   #r := FALSE;
   #a1 := W#16#0000;
   #a2 := W#16#0000;
   #activeDataBlock := 0;
   // PB4, STEP 5 network 1
   #a2 := #a1;
   #a1 := "ROLL_GetM"(FirstByte := 239, Width := 8);
   #a2 := #a1;
   #a1 := W#16#001E;
   #comparisonResults[0] := (WORD_TO_INT(#a2) = WORD_TO_INT(#a1));
   #r := #comparisonResults[0];
   "ROLL_State".M[23, 5] := #r;
   // PB4, STEP 5 network 2
   #a2 := #a1;
   #a1 := "ROLL_GetM"(FirstByte := 239, Width := 8);
   #a2 := #a1;
   #a1 := W#16#001F;
   #comparisonResults[1] := (WORD_TO_INT(#a2) = WORD_TO_INT(#a1));
   #r := #comparisonResults[1];
   "ROLL_State".M[23, 6] := #r;
   // PB4, STEP 5 network 3
   #a2 := #a1;
   #a1 := "ROLL_GetM"(FirstByte := 239, Width := 8);
   #a2 := #a1;
   #a1 := W#16#0023;
   #comparisonResults[2] := (WORD_TO_INT(#a2) = WORD_TO_INT(#a1));
   #r := #comparisonResults[2];
   "ROLL_State".M[24, 0] := #r;
   // PB4, STEP 5 network 4
   #a2 := #a1;
   #a1 := "ROLL_GetM"(FirstByte := 239, Width := 8);
   #a2 := #a1;
   #a1 := W#16#0024;
   #comparisonResults[3] := (WORD_TO_INT(#a2) = WORD_TO_INT(#a1));
   #r := #comparisonResults[3];
   "ROLL_State".M[24, 1] := #r;
   // PB4, STEP 5 network 5
   #a2 := #a1;
   #a1 := "ROLL_GetM"(FirstByte := 239, Width := 8);
   #a2 := #a1;
   #a1 := W#16#0025;
   #comparisonResults[4] := (WORD_TO_INT(#a2) = WORD_TO_INT(#a1));
   #r := #comparisonResults[4];
   "ROLL_State".M[24, 2] := #r;
   // PB4, STEP 5 network 6
   #a2 := #a1;
   #a1 := "ROLL_GetM"(FirstByte := 239, Width := 8);
   #a2 := #a1;
   #a1 := W#16#0026;
   #comparisonResults[5] := (WORD_TO_INT(#a2) = WORD_TO_INT(#a1));
   #r := #comparisonResults[5];
   "ROLL_State".M[24, 3] := #r;
   // PB4, STEP 5 network 7
   #a2 := #a1;
   #a1 := "ROLL_GetM"(FirstByte := 239, Width := 8);
   #a2 := #a1;
   #a1 := W#16#0027;
   #comparisonResults[6] := (WORD_TO_INT(#a2) = WORD_TO_INT(#a1));
   #r := #comparisonResults[6];
   "ROLL_State".M[24, 4] := #r;
   // PB4, STEP 5 network 8
   #a2 := #a1;
   #a1 := "ROLL_GetM"(FirstByte := 239, Width := 8);
   #a2 := #a1;
   #a1 := W#16#0032;
   #comparisonResults[7] := (WORD_TO_INT(#a2) = WORD_TO_INT(#a1));
   #r := #comparisonResults[7];
   "ROLL_State".M[25, 0] := #r;
   // PB4, STEP 5 network 9
   #a2 := #a1;
   #a1 := "ROLL_GetM"(FirstByte := 239, Width := 8);
   #a2 := #a1;
   #a1 := W#16#0033;
   #comparisonResults[8] := (WORD_TO_INT(#a2) = WORD_TO_INT(#a1));
   #r := #comparisonResults[8];
   "ROLL_State".M[25, 1] := #r;
   // PB4, STEP 5 network 10
   #a2 := #a1;
   #a1 := "ROLL_GetM"(FirstByte := 239, Width := 8);
   #a2 := #a1;
   #a1 := W#16#0034;
   #comparisonResults[9] := (WORD_TO_INT(#a2) = WORD_TO_INT(#a1));
   #r := #comparisonResults[9];
   "ROLL_State".M[25, 2] := #r;
   // PB4, STEP 5 network 11
   #a2 := #a1;
   #a1 := "ROLL_GetM"(FirstByte := 239, Width := 8);
   #a2 := #a1;
   #a1 := W#16#0035;
   #comparisonResults[10] := (WORD_TO_INT(#a2) = WORD_TO_INT(#a1));
   #r := #comparisonResults[10];
   "ROLL_State".M[25, 3] := #r;
   // PB4, STEP 5 network 12
   #a2 := #a1;
   #a1 := "ROLL_GetM"(FirstByte := 239, Width := 8);
   #a2 := #a1;
   #a1 := W#16#0037;
   #comparisonResults[11] := (WORD_TO_INT(#a2) = WORD_TO_INT(#a1));
   #r := #comparisonResults[11];
   "ROLL_State".M[25, 4] := #r;
   // PB4, STEP 5 network 13
   #a2 := #a1;
   #a1 := "ROLL_GetM"(FirstByte := 239, Width := 8);
   #a2 := #a1;
   #a1 := W#16#0038;
   #comparisonResults[12] := (WORD_TO_INT(#a2) = WORD_TO_INT(#a1));
   #r := #comparisonResults[12];
   "ROLL_State".M[25, 5] := #r;
   // PB4, STEP 5 network 14
   #a2 := #a1;
   #a1 := "ROLL_GetM"(FirstByte := 239, Width := 8);
   #a2 := #a1;
   #a1 := W#16#0039;
   #comparisonResults[13] := (WORD_TO_INT(#a2) = WORD_TO_INT(#a1));
   #r := #comparisonResults[13];
   "ROLL_State".M[25, 6] := #r;
   // PB4, STEP 5 network 15
   #a2 := #a1;
   #a1 := "ROLL_GetM"(FirstByte := 239, Width := 8);
   #a2 := #a1;
   #a1 := W#16#003A;
   #comparisonResults[14] := (WORD_TO_INT(#a2) = WORD_TO_INT(#a1));
   #r := #comparisonResults[14];
   "ROLL_State".M[25, 7] := #r;
   // PB4, STEP 5 network 16
   #a2 := #a1;
   #a1 := "ROLL_GetM"(FirstByte := 239, Width := 8);
   #a2 := #a1;
   #a1 := W#16#003C;
   #comparisonResults[15] := (WORD_TO_INT(#a2) = WORD_TO_INT(#a1));
   #r := #comparisonResults[15];
   "ROLL_State".M[26, 0] := #r;
   // PB4, STEP 5 network 17
   #a2 := #a1;
   #a1 := "ROLL_GetM"(FirstByte := 239, Width := 8);
   #a2 := #a1;
   #a1 := W#16#003D;
   #comparisonResults[16] := (WORD_TO_INT(#a2) = WORD_TO_INT(#a1));
   #r := #comparisonResults[16];
   "ROLL_State".M[26, 1] := #r;
   // PB4, STEP 5 network 18
   #a2 := #a1;
   #a1 := "ROLL_GetM"(FirstByte := 239, Width := 8);
   #a2 := #a1;
   #a1 := W#16#003E;
   #comparisonResults[17] := (WORD_TO_INT(#a2) = WORD_TO_INT(#a1));
   #r := #comparisonResults[17];
   "ROLL_State".M[26, 2] := #r;
   // PB4, STEP 5 network 19
   #a2 := #a1;
   #a1 := "ROLL_GetM"(FirstByte := 239, Width := 8);
   #a2 := #a1;
   #a1 := W#16#003F;
   #comparisonResults[18] := (WORD_TO_INT(#a2) = WORD_TO_INT(#a1));
   #r := #comparisonResults[18];
   "ROLL_State".M[26, 3] := #r;
   // PB4, STEP 5 network 20
   #a2 := #a1;
   #a1 := "ROLL_GetM"(FirstByte := 239, Width := 8);
   #a2 := #a1;
   #a1 := W#16#0041;
   #comparisonResults[19] := (WORD_TO_INT(#a2) = WORD_TO_INT(#a1));
   #r := #comparisonResults[19];
   "ROLL_State".M[26, 5] := #r;
   // PB4, STEP 5 network 21
   #a2 := #a1;
   #a1 := "ROLL_GetM"(FirstByte := 239, Width := 8);
   #a2 := #a1;
   #a1 := W#16#0042;
   #comparisonResults[20] := (WORD_TO_INT(#a2) = WORD_TO_INT(#a1));
   #r := #comparisonResults[20];
   "ROLL_State".M[26, 6] := #r;
   // PB4, STEP 5 network 22
   #a2 := #a1;
   #a1 := "ROLL_GetM"(FirstByte := 239, Width := 8);
   #a2 := #a1;
   #a1 := W#16#0045;
   #comparisonResults[21] := (WORD_TO_INT(#a2) = WORD_TO_INT(#a1));
   #r := #comparisonResults[21];
   "ROLL_State".M[27, 1] := #r;
   // PB4, STEP 5 network 23
   #a2 := #a1;
   #a1 := "ROLL_GetM"(FirstByte := 239, Width := 8);
   #a2 := #a1;
   #a1 := W#16#0048;
   #comparisonResults[22] := (WORD_TO_INT(#a2) = WORD_TO_INT(#a1));
   #r := #comparisonResults[22];
   "ROLL_State".M[27, 4] := #r;
   // PB4, STEP 5 network 24
   #a2 := #a1;
   #a1 := "ROLL_GetM"(FirstByte := 239, Width := 8);
   #a2 := #a1;
   #a1 := W#16#0049;
   #comparisonResults[23] := (WORD_TO_INT(#a2) = WORD_TO_INT(#a1));
   #r := #comparisonResults[23];
   "ROLL_State".M[27, 5] := #r;
   // PB4, STEP 5 network 25
   #a2 := #a1;
   #a1 := "ROLL_GetM"(FirstByte := 239, Width := 8);
   #a2 := #a1;
   #a1 := W#16#0063;
   #comparisonResults[24] := (WORD_TO_INT(#a2) = WORD_TO_INT(#a1));
   #r := #comparisonResults[24];
   "ROLL_State".M[27, 7] := #r;
   // PB4, STEP 5 network 26
   RETURN;
END_FUNCTION

FUNCTION "ROLL_PB50" : Void   // FC33, SCL
{ S7_Optimized_Access := 'TRUE' }
VERSION : 0.1
// stored: AutoNumber true, IsIECCheckEnabled false, SetENOAutomatically false, UDAEnableTagReadback false
   VAR_TEMP
      r : Bool;
      a1 : Word;
      a2 : Word;
      activeDataBlock : Int;
      comparisonResults : Array[0..0] of Bool;
   END_VAR
BEGIN

   #r := FALSE;
   #a1 := W#16#0000;
   #a2 := W#16#0000;
   #activeDataBlock := 0;
   // PB50, STEP 5 network 1
   #activeDataBlock := 15;
   // PB50, STEP 5 network 2
   #r := "ROLL_State".M[0, 1];
   IF #r THEN
       "ROLL_State".M[0, 2] := FALSE;
   END_IF;
   // PB50, STEP 5 network 3
   #a2 := #a1;
   #a1 := W#16#2008;
   #r := ((NOT "ROLL_State".M[0, 1]) AND "ROLL_IO".Input[3, 0]);
   "ROLL_TimerOp"(Number := 11,
                  Operation := 0,
                  Signal := #r,
                  Preset := #a1);
   // PB50, STEP 5 network 4
   #a2 := #a1;
   #a1 := W#16#1020;
   #r := "ROLL_State".M[29, 0];
   "ROLL_TimerOp"(Number := 13,
                  Operation := 0,
                  Signal := #r,
                  Preset := #a1);
   // PB50, STEP 5 network 5
   RETURN;
END_FUNCTION

FUNCTION "ROLL_PB51" : Void   // FC34, SCL
{ S7_Optimized_Access := 'TRUE' }
VERSION : 0.1
// stored: AutoNumber true, IsIECCheckEnabled false, SetENOAutomatically false, UDAEnableTagReadback false
   VAR_TEMP
      r : Bool;
      a1 : Word;
      a2 : Word;
      activeDataBlock : Int;
      comparisonResults : Array[0..0] of Bool;
   END_VAR
BEGIN

   #r := FALSE;
   #a1 := W#16#0000;
   #a2 := W#16#0000;
   #activeDataBlock := 0;
   // PB51, STEP 5 network 1
   #a2 := #a1;
   #a1 := W#16#2060;
   #r := "ROLL_IO".Output[24, 0];
   "ROLL_TimerOp"(Number := 15,
                  Operation := 0,
                  Signal := #r,
                  Preset := #a1);
   // PB51, STEP 5 network 2
   #a2 := #a1;
   #a1 := W#16#3360;
   #r := ((NOT "ROLL_IO".Input[5, 6]) AND "ROLL_State".M[31, 5]);
   "ROLL_TimerOp"(Number := 16,
                  Operation := 0,
                  Signal := #r,
                  Preset := #a1);
   // PB51, STEP 5 network 3
   #a2 := #a1;
   #a1 := W#16#1010;
   #r := "ROLL_State".M[37, 5];
   "ROLL_TimerOp"(Number := 18,
                  Operation := 0,
                  Signal := #r,
                  Preset := #a1);
   // PB51, STEP 5 network 4
   #a2 := #a1;
   #a1 := W#16#2015;
   #r := (((NOT "ROLL_IO".Input[124, 1]) AND "ROLL_IO".Output[112, 1]) OR ((NOT "ROLL_IO".Input[124, 2]) AND "ROLL_IO".Output[112, 2]));
   "ROLL_TimerOp"(Number := 19,
                  Operation := 0,
                  Signal := #r,
                  Preset := #a1);
   // PB51, STEP 5 network 5
   #a2 := #a1;
   #a1 := W#16#1010;
   #r := (("ROLL_IO".Input[123, 4] OR "ROLL_IO".Input[123, 5]) AND "ROLL_IO".Output[112, 0]);
   "ROLL_TimerOp"(Number := 20,
                  Operation := 0,
                  Signal := #r,
                  Preset := #a1);
   // PB51, STEP 5 network 6
   #a2 := #a1;
   #a1 := W#16#1050;
   #r := "ROLL_IO".Input[123, 4];
   "ROLL_TimerOp"(Number := 21,
                  Operation := 0,
                  Signal := #r,
                  Preset := #a1);
   // PB51, STEP 5 network 7
   #a2 := #a1;
   #a1 := W#16#2005;
   #r := ("ROLL_IO".Input[125, 0] AND "ROLL_IO".Input[125, 1]);
   "ROLL_TimerOp"(Number := 95,
                  Operation := 0,
                  Signal := #r,
                  Preset := #a1);
   // PB51, STEP 5 network 8
   RETURN;
END_FUNCTION

FUNCTION "ROLL_PB52" : Void   // FC35, SCL
{ S7_Optimized_Access := 'TRUE' }
VERSION : 0.1
// stored: AutoNumber true, IsIECCheckEnabled false, SetENOAutomatically false, UDAEnableTagReadback false
   VAR_TEMP
      r : Bool;
      a1 : Word;
      a2 : Word;
      activeDataBlock : Int;
      comparisonResults : Array[0..0] of Bool;
   END_VAR
BEGIN

   #r := FALSE;
   #a1 := W#16#0000;
   #a2 := W#16#0000;
   #activeDataBlock := 0;
   // PB52, STEP 5 network 1
   #activeDataBlock := 15;
   // PB52, STEP 5 network 2
   #a2 := #a1;
   #a1 := "ROLL_GetDW"(DbNumber := #activeDataBlock, Index := 17);
   #r := ((NOT "ROLL_IO".Input[5, 5]) AND (NOT "ROLL_State".M[6, 3]) AND "ROLL_IO".Input[3, 1] AND "ROLL_State".M[4, 1] AND "ROLL_State".M[40, 5]);
   "ROLL_TimerOp"(Number := 17,
                  Operation := 0,
                  Signal := #r,
                  Preset := #a1);
   // PB52, STEP 5 network 3
   #a2 := #a1;
   #a1 := "ROLL_GetDW"(DbNumber := #activeDataBlock, Index := 31);
   #r := ((NOT "ROLL_IO".Input[5, 3]) AND (NOT "ROLL_State".M[6, 1]) AND "ROLL_IO".Input[3, 1] AND "ROLL_State".M[4, 1]);
   "ROLL_TimerOp"(Number := 31,
                  Operation := 0,
                  Signal := #r,
                  Preset := #a1);
   // PB52, STEP 5 network 4
   #a2 := #a1;
   #a1 := "ROLL_GetDW"(DbNumber := #activeDataBlock, Index := 32);
   #r := ((NOT "ROLL_IO".Input[6, 0]) AND (NOT "ROLL_State".M[6, 4]) AND "ROLL_IO".Input[3, 1] AND "ROLL_State".M[4, 1]);
   "ROLL_TimerOp"(Number := 32,
                  Operation := 0,
                  Signal := #r,
                  Preset := #a1);
   // PB52, STEP 5 network 5
   #a2 := #a1;
   #a1 := "ROLL_GetDW"(DbNumber := #activeDataBlock, Index := 33);
   #r := ((NOT "ROLL_IO".Input[6, 2]) AND (NOT "ROLL_State".M[6, 5]) AND "ROLL_IO".Input[3, 1] AND "ROLL_State".M[4, 1]);
   "ROLL_TimerOp"(Number := 33,
                  Operation := 0,
                  Signal := #r,
                  Preset := #a1);
   // PB52, STEP 5 network 6
   #a2 := #a1;
   #a1 := W#16#3030;
   #r := ((NOT "ROLL_State".M[0, 4]) AND (NOT "ROLL_State".M[6, 7]) AND "ROLL_IO".Input[3, 1] AND "ROLL_State".M[4, 1]);
   "ROLL_TimerOp"(Number := 35,
                  Operation := 0,
                  Signal := #r,
                  Preset := #a1);
   // PB52, STEP 5 network 7
   #a2 := #a1;
   #a1 := W#16#3030;
   #r := ((NOT "ROLL_State".M[0, 4]) AND (NOT "ROLL_State".M[7, 0]) AND "ROLL_IO".Input[3, 1] AND "ROLL_State".M[4, 1]);
   "ROLL_TimerOp"(Number := 36,
                  Operation := 0,
                  Signal := #r,
                  Preset := #a1);
   // PB52, STEP 5 network 8
   #a2 := #a1;
   #a1 := W#16#3030;
   #r := ((NOT "ROLL_State".M[0, 4]) AND (NOT "ROLL_State".M[7, 1]) AND "ROLL_IO".Input[3, 1] AND "ROLL_State".M[4, 1]);
   "ROLL_TimerOp"(Number := 37,
                  Operation := 0,
                  Signal := #r,
                  Preset := #a1);
   // PB52, STEP 5 network 9
   #a2 := #a1;
   #a1 := W#16#3030;
   #r := ((NOT "ROLL_State".M[0, 4]) AND (NOT "ROLL_State".M[7, 2]) AND "ROLL_IO".Input[3, 1] AND "ROLL_State".M[4, 1]);
   "ROLL_TimerOp"(Number := 38,
                  Operation := 0,
                  Signal := #r,
                  Preset := #a1);
   // PB52, STEP 5 network 10
   #a2 := #a1;
   #a1 := W#16#1005;
   #r := "ROLL_IO".Input[123, 1];
   "ROLL_TimerOp"(Number := 45,
                  Operation := 0,
                  Signal := #r,
                  Preset := #a1);
   // PB52, STEP 5 network 11
   #a2 := #a1;
   #a1 := "ROLL_GetDW"(DbNumber := #activeDataBlock, Index := 58);
   #r := ("ROLL_IO".Input[3, 1] AND "ROLL_State".M[3, 6]);
   "ROLL_TimerOp"(Number := 58,
                  Operation := 1,
                  Signal := #r,
                  Preset := #a1);
   #a2 := #a1;
   #a1 := "ROLL_GetDW"(DbNumber := #activeDataBlock, Index := 59);
   #r := ("ROLL_State".M[3, 6] AND "ROLL_State".S5Timers[58].Q);
   "ROLL_TimerOp"(Number := 59,
                  Operation := 1,
                  Signal := #r,
                  Preset := #a1);
   // PB52, STEP 5 network 12
   #a2 := #a1;
   #a1 := "ROLL_GetDW"(DbNumber := #activeDataBlock, Index := 63);
   #r := (NOT "ROLL_State".S5Timers[62].Q);
   "ROLL_TimerOp"(Number := 63,
                  Operation := 0,
                  Signal := #r,
                  Preset := #a1);
   #a2 := #a1;
   #a1 := "ROLL_GetDW"(DbNumber := #activeDataBlock, Index := 62);
   #r := "ROLL_State".S5Timers[63].Q;
   "ROLL_TimerOp"(Number := 62,
                  Operation := 1,
                  Signal := #r,
                  Preset := #a1);
   #r := ((NOT "ROLL_State".M[103, 0]) AND (NOT "ROLL_State".M[103, 3]) AND (NOT "ROLL_State".M[103, 4]) AND (NOT "ROLL_State".S5Timers[119].Q));
   "ROLL_TimerOp"(Number := 62,
                  Operation := 2,
                  Signal := #r,
                  Preset := #a1);
   // PB52, STEP 5 network 13
   #a2 := #a1;
   #a1 := W#16#2010;
   #r := "ROLL_IO".Input[5, 3];
   "ROLL_TimerOp"(Number := 70,
                  Operation := 1,
                  Signal := #r,
                  Preset := #a1);
   // PB52, STEP 5 network 14
   #a2 := #a1;
   #a1 := W#16#2010;
   #r := "ROLL_IO".Input[6, 2];
   "ROLL_TimerOp"(Number := 72,
                  Operation := 1,
                  Signal := #r,
                  Preset := #a1);
   // PB52, STEP 5 network 15
   #a2 := #a1;
   #a1 := "ROLL_GetDW"(DbNumber := #activeDataBlock, Index := 85);
   #r := "ROLL_State".M[41, 0];
   "ROLL_TimerOp"(Number := 85,
                  Operation := 1,
                  Signal := #r,
                  Preset := #a1);
   // PB52, STEP 5 network 16
   RETURN;
END_FUNCTION

FUNCTION "ROLL_PB7" : Void   // FC17, SCL
{ S7_Optimized_Access := 'TRUE' }
VERSION : 0.1
// stored: AutoNumber true, IsIECCheckEnabled false, SetENOAutomatically false, UDAEnableTagReadback false
   VAR_TEMP
      r : Bool;
      a1 : Word;
      a2 : Word;
      activeDataBlock : Int;
      comparisonResults : Array[0..0] of Bool;
   END_VAR
BEGIN

   #r := FALSE;
   #a1 := W#16#0000;
   #a2 := W#16#0000;
   #activeDataBlock := 0;
   // PB7, STEP 5 network 1
   #r := ((NOT "ROLL_State".M[70, 2]) AND (NOT "ROLL_State".M[70, 3]) AND (NOT "ROLL_State".M[70, 4]) AND (NOT "ROLL_State".M[70, 6]) AND "ROLL_IO".Input[11, 0] AND "ROLL_IO".Input[11, 6] AND "ROLL_IO".Input[13, 3] AND "ROLL_State".M[63, 1]);
   "ROLL_State".M[28, 0] := #r;
   // PB7, STEP 5 network 2
   #r := ("ROLL_IO".Input[12, 1] AND "ROLL_IO".Input[12, 7]);
   "ROLL_State".M[28, 1] := #r;
   // PB7, STEP 5 network 3
   #r := ((NOT "ROLL_IO".Output[112, 5]) AND ((NOT "ROLL_IO".Output[112, 0]) OR (NOT "ROLL_State".M[31, 4])));
   "ROLL_State".M[28, 2] := #r;
   // PB7, STEP 5 network 4
   #r := (((NOT "ROLL_IO".Output[113, 0]) AND (NOT "ROLL_IO".Output[113, 1]) AND (NOT "ROLL_IO".Output[113, 3]) AND (NOT "ROLL_IO".Output[113, 5]) AND (NOT "ROLL_IO".Input[123, 5]) AND (NOT "ROLL_IO".Input[123, 6]) AND "ROLL_IO".Output[113, 2] AND "ROLL_IO".Output[113, 4] AND "ROLL_IO".Input[124, 1] AND "ROLL_IO".Input[124, 4]) OR "ROLL_State".M[0, 4]);
   "ROLL_State".M[240, 0] := #r;
   // PB7, STEP 5 network 5
   #r := ((((NOT "ROLL_IO".Output[113, 2]) AND "ROLL_IO".Output[113, 3] AND "ROLL_IO".Input[123, 5] AND "ROLL_IO".Input[124, 1] AND "ROLL_IO".Input[124, 4]) OR ((NOT "ROLL_IO".Output[113, 3]) AND "ROLL_IO".Output[113, 2] AND "ROLL_IO".Input[124, 1] AND "ROLL_IO".Input[124, 5]) OR "ROLL_State".M[0, 4]) AND "ROLL_State".M[20, 2]);
   "ROLL_State".M[240, 1] := #r;
   // PB7, STEP 5 network 6
   #r := ("ROLL_State".M[240, 0] OR "ROLL_State".M[240, 1]);
   "ROLL_State".M[28, 3] := #r;
   // PB7, STEP 5 network 7
   #r := ("ROLL_State".M[28, 0] AND "ROLL_State".M[28, 1] AND "ROLL_State".M[28, 2] AND "ROLL_State".M[28, 3]);
   "ROLL_State".M[28, 4] := #r;
   // PB7, STEP 5 network 8
   #r := ("ROLL_IO".Input[10, 7] AND "ROLL_IO".Input[3, 4] AND "ROLL_IO".Input[3, 5] AND "ROLL_IO".Input[3, 7]);
   "ROLL_State".M[28, 5] := #r;
   // PB7, STEP 5 network 9
   #r := ((NOT "ROLL_State".M[13, 4]) AND (NOT "ROLL_State".M[16, 6]) AND (NOT "ROLL_State".M[5, 7]) AND "ROLL_State".M[28, 5]);
   "ROLL_State".M[28, 6] := #r;
   // PB7, STEP 5 network 10
   #r := (("ROLL_IO".Input[0, 2] AND "ROLL_IO".Input[0, 4]) OR "ROLL_IO".Input[0, 1]);
   IF #r THEN
       "ROLL_State".M[29, 0] := TRUE;
   END_IF;
   #r := (NOT "ROLL_State".M[28, 6]);
   IF #r THEN
       "ROLL_State".M[29, 0] := FALSE;
   END_IF;
   // PB7, STEP 5 network 11
   #r := ("ROLL_State".M[29, 0] AND "ROLL_State".S5Timers[13].Q);
   "ROLL_State".M[29, 1] := #r;
   // PB7, STEP 5 network 12
   #r := (NOT "ROLL_State".M[12, 1]);
   "ROLL_State".M[30, 0] := #r;
   // PB7, STEP 5 network 13
   #r := "ROLL_State".M[0, 4];
   "ROLL_State".M[30, 1] := #r;
   // PB7, STEP 5 network 14
   #r := ((NOT "ROLL_State".M[6, 1]) AND (NOT "ROLL_State".M[6, 3]) AND (NOT "ROLL_State".M[6, 4]) AND (NOT "ROLL_State".M[6, 5]) AND (NOT "ROLL_State".M[6, 6]) AND (NOT "ROLL_State".M[6, 7]) AND (NOT "ROLL_State".M[7, 0]) AND (NOT "ROLL_State".M[7, 1]) AND (NOT "ROLL_State".M[7, 2]) AND (NOT "ROLL_State".M[7, 3]) AND (NOT "ROLL_State".M[7, 7]));
   "ROLL_State".M[30, 2] := #r;
   // PB7, STEP 5 network 15
   #r := ((NOT "ROLL_IO".Input[3, 6]) AND (NOT "ROLL_State".M[5, 6]));
   "ROLL_State".M[30, 3] := #r;
   // PB7, STEP 5 network 16
   #r := (("ROLL_State".M[30, 0] AND "ROLL_State".M[30, 1] AND "ROLL_State".M[30, 2] AND "ROLL_State".M[30, 3]) OR "ROLL_IO".Input[0, 0] OR "ROLL_IO".Input[0, 6]);
   "ROLL_State".M[30, 5] := #r;
   // PB7, STEP 5 network 17
   #r := ((NOT "ROLL_State".M[11, 0]) AND (NOT "ROLL_State".M[13, 1]) AND (NOT "ROLL_State".M[13, 3]) AND (NOT "ROLL_State".M[5, 0]) AND (NOT "ROLL_State".M[5, 1]) AND (NOT "ROLL_State".M[5, 2]));
   "ROLL_State".M[30, 6] := #r;
   // PB7, STEP 5 network 18
   #r := ((NOT "ROLL_State".M[11, 1]) AND (NOT "ROLL_State".M[5, 3]) AND (NOT "ROLL_State".M[9, 1]) AND (NOT "ROLL_State".M[9, 2]) AND (NOT "ROLL_State".M[9, 3]) AND "ROLL_IO".Input[8, 5] AND "ROLL_State".M[28, 6]);
   "ROLL_State".M[30, 7] := #r;
   // PB7, STEP 5 network 19
   #r := ((NOT "ROLL_State".M[12, 0]) AND (NOT "ROLL_State".M[9, 0]));
   "ROLL_State".M[31, 0] := #r;
   // PB7, STEP 5 network 20
   #r := ((NOT "ROLL_State".M[87, 5]) AND (NOT "ROLL_State".M[88, 1]) AND (NOT "ROLL_State".M[88, 3]) AND (NOT "ROLL_State".M[88, 4]) AND (NOT "ROLL_State".M[88, 5]) AND (NOT "ROLL_State".M[88, 6]));
   "ROLL_State".M[31, 2] := #r;
   // PB7, STEP 5 network 21
   #r := ("ROLL_State".M[30, 5] AND "ROLL_State".M[30, 6] AND "ROLL_State".M[30, 7] AND "ROLL_State".M[31, 0] AND "ROLL_State".M[31, 2]);
   "ROLL_State".M[31, 1] := #r;
   // PB7, STEP 5 network 22
   #r := (("ROLL_State".M[28, 4] OR "ROLL_State".M[31, 5]) AND "ROLL_IO".Input[0, 4] AND "ROLL_State".M[4, 4]);
   IF #r THEN
       "ROLL_State".M[31, 4] := TRUE;
   END_IF;
   #r := ((NOT "ROLL_IO".Input[0, 2]) OR (NOT "ROLL_IO".Input[0, 3]) OR (NOT "ROLL_State".M[29, 0]) OR (NOT "ROLL_State".M[31, 1]));
   IF #r THEN
       "ROLL_State".M[31, 4] := FALSE;
   END_IF;
   // PB7, STEP 5 network 23
   #r := "ROLL_State".M[31, 4];
   IF #r THEN
       "ROLL_State".M[31, 5] := TRUE;
   END_IF;
   #r := (((NOT "ROLL_State".M[31, 4]) AND (((NOT "ROLL_State".M[37, 2]) AND "ROLL_State".M[37, 1]) OR "ROLL_State".M[37, 0]) AND "ROLL_State".M[28, 4]) OR (NOT "ROLL_IO".Input[0, 2]));
   IF #r THEN
       "ROLL_State".M[31, 5] := FALSE;
   END_IF;
   // PB7, STEP 5 network 24
   #r := "ROLL_State".M[52, 3];
   IF #r THEN
       "ROLL_State".M[31, 6] := TRUE;
   END_IF;
   #r := ((NOT "ROLL_IO".Input[14, 0]) AND "ROLL_IO".Input[12, 1]);
   IF #r THEN
       "ROLL_State".M[31, 6] := FALSE;
   END_IF;
   // PB7, STEP 5 network 25
   #r := "ROLL_State".M[31, 5];
   "ROLL_IO".Output[16, 6] := #r;
   // PB7, STEP 5 network 26
   #r := "ROLL_State".M[40, 0];
   "ROLL_IO".Output[16, 7] := #r;
   // PB7, STEP 5 network 27
   RETURN;
END_FUNCTION

FUNCTION "ROLL_PB8" : Void   // FC18, SCL
{ S7_Optimized_Access := 'TRUE' }
VERSION : 0.1
// stored: AutoNumber true, IsIECCheckEnabled false, SetENOAutomatically false, UDAEnableTagReadback false
   VAR_TEMP
      r : Bool;
      a1 : Word;
      a2 : Word;
      activeDataBlock : Int;
      comparisonResults : Array[0..0] of Bool;
   END_VAR
BEGIN

   #r := FALSE;
   #a1 := W#16#0000;
   #a2 := W#16#0000;
   #activeDataBlock := 0;
   // PB8, STEP 5 network 1
   #r := ("ROLL_State".M[37, 7] OR "ROLL_State".M[38, 0] OR "ROLL_State".M[39, 7] OR "ROLL_State".M[40, 0] OR "ROLL_State".M[40, 1] OR "ROLL_State".M[40, 4] OR "ROLL_State".M[41, 0] OR "ROLL_State".M[41, 6] OR "ROLL_State".M[41, 7] OR "ROLL_State".M[42, 2] OR "ROLL_State".M[42, 3]);
   "ROLL_State".M[33, 0] := #r;
   // PB8, STEP 5 network 2
   #r := (((NOT "ROLL_State".M[16, 0]) AND (NOT "ROLL_State".M[16, 1]) AND (NOT "ROLL_State".M[16, 4]) AND "ROLL_State".M[37, 2]) OR "ROLL_State".M[37, 3] OR "ROLL_State".M[37, 5] OR "ROLL_State".M[37, 6] OR "ROLL_State".M[39, 4] OR "ROLL_State".M[39, 5] OR "ROLL_State".M[40, 2] OR "ROLL_State".M[40, 3] OR "ROLL_State".M[40, 6] OR "ROLL_State".M[40, 7] OR "ROLL_State".M[41, 2] OR "ROLL_State".M[42, 0] OR "ROLL_State".M[42, 4]);
   "ROLL_State".M[33, 1] := #r;
   // PB8, STEP 5 network 3
   #a2 := #a1;
   #a1 := W#16#2030;
   #r := ((NOT "ROLL_State".M[3, 1]) AND ("ROLL_State".M[33, 0] OR "ROLL_State".M[42, 6] OR "ROLL_State".M[43, 4] OR "ROLL_State".M[43, 6] OR "ROLL_State".M[43, 7] OR "ROLL_State".M[44, 2] OR "ROLL_State".M[45, 0] OR "ROLL_State".M[45, 1] OR "ROLL_State".M[45, 5] OR "ROLL_State".M[45, 7] OR "ROLL_State".M[46, 1] OR "ROLL_State".M[46, 4] OR "ROLL_State".M[46, 6] OR "ROLL_State".M[52, 1] OR "ROLL_State".M[52, 2] OR "ROLL_State".M[53, 3]) AND "ROLL_IO".Input[0, 2] AND "ROLL_State".M[29, 0]);
   "ROLL_TimerOp"(Number := 40,
                  Operation := 0,
                  Signal := #r,
                  Preset := #a1);
   // PB8, STEP 5 network 4
   #a2 := #a1;
   #a1 := W#16#2030;
   #r := ((NOT "ROLL_State".M[3, 1]) AND (((NOT "ROLL_IO".Input[11, 2]) AND "ROLL_State".M[52, 0]) OR ((NOT "ROLL_State".M[15, 1]) AND "ROLL_State".M[53, 1]) OR "ROLL_State".M[33, 1] OR "ROLL_State".M[43, 0] OR "ROLL_State".M[43, 2] OR "ROLL_State".M[43, 3] OR "ROLL_State".M[44, 0] OR "ROLL_State".M[44, 7] OR "ROLL_State".M[45, 3] OR "ROLL_State".M[45, 4] OR "ROLL_State".M[46, 2] OR "ROLL_State".M[46, 3] OR "ROLL_State".M[46, 7] OR "ROLL_State".M[47, 3] OR "ROLL_State".M[52, 3] OR "ROLL_State".M[53, 2] OR "ROLL_State".M[53, 5] OR "ROLL_State".M[53, 6]) AND "ROLL_IO".Input[0, 2] AND "ROLL_State".M[29, 0]);
   "ROLL_TimerOp"(Number := 41,
                  Operation := 0,
                  Signal := #r,
                  Preset := #a1);
   // PB8, STEP 5 network 5
   #r := ("ROLL_State".S5Timers[40].Q OR "ROLL_State".S5Timers[41].Q);
   IF #r THEN
       "ROLL_State".M[34, 1] := TRUE;
   END_IF;
   #r := ((NOT "ROLL_IO".Input[0, 2]) OR "ROLL_State".M[3, 1]);
   IF #r THEN
       "ROLL_State".M[34, 1] := FALSE;
   END_IF;
   // PB8, STEP 5 network 6
   RETURN;
END_FUNCTION

FUNCTION "ROLL_PB9" : Void   // FC19, SCL
{ S7_Optimized_Access := 'TRUE' }
VERSION : 0.1
// stored: AutoNumber true, IsIECCheckEnabled false, SetENOAutomatically false, UDAEnableTagReadback false
   VAR_TEMP
      r : Bool;
      a1 : Word;
      a2 : Word;
      activeDataBlock : Int;
      comparisonResults : Array[0..0] of Bool;
   END_VAR
BEGIN

   #r := FALSE;
   #a1 := W#16#0000;
   #a2 := W#16#0000;
   #activeDataBlock := 0;
   // PB9, STEP 5 network 1
   #r := ((NOT "ROLL_State".M[32, 1]) AND (NOT "ROLL_State".M[32, 2]) AND "ROLL_IO".Input[0, 2]);
   "ROLL_State".M[32, 0] := #r;
   // PB9, STEP 5 network 2
   #r := "ROLL_State".M[32, 0];
   IF #r THEN
       "ROLL_State".M[32, 1] := TRUE;
   END_IF;
   #r := ((NOT "ROLL_IO".Input[0, 2]) OR "ROLL_IO".Input[0, 1] OR "ROLL_State".M[32, 2]);
   IF #r THEN
       "ROLL_State".M[32, 1] := FALSE;
   END_IF;
   // PB9, STEP 5 network 3
   #r := ((NOT "ROLL_IO".Input[0, 2]) OR "ROLL_IO".Input[0, 1]);
   "ROLL_State".M[32, 2] := #r;
   // PB9, STEP 5 network 4
   #r := ((NOT "ROLL_State".M[12, 0]) AND (NOT "ROLL_State".M[5, 0]) AND (NOT "ROLL_State".M[5, 2]) AND (NOT "ROLL_State".M[9, 0]));
   "ROLL_State".M[35, 1] := #r;
   // PB9, STEP 5 network 5
   #r := "ROLL_IO".Input[0, 4];
   IF #r THEN
       "ROLL_State".M[35, 2] := TRUE;
   END_IF;
   #r := ((NOT "ROLL_State".M[29, 0]) OR (NOT "ROLL_State".M[31, 5]) OR (NOT "ROLL_State".M[35, 1]) OR "ROLL_State".M[16, 3]);
   IF #r THEN
       "ROLL_State".M[35, 2] := FALSE;
   END_IF;
   // PB9, STEP 5 network 6
   #r := ("ROLL_State".M[32, 0] OR "ROLL_State".M[53, 6]);
   IF #r THEN
       "ROLL_State".M[37, 0] := TRUE;
   END_IF;
   #r := ("ROLL_State".M[32, 2] OR "ROLL_State".M[37, 1] OR "ROLL_State".M[38, 0] OR "ROLL_State".M[39, 5]);
   IF #r THEN
       "ROLL_State".M[37, 0] := FALSE;
   END_IF;
   // PB9, STEP 5 network 7
   #r := ((NOT "ROLL_IO".Input[123, 5]) AND (NOT "ROLL_IO".Input[123, 6]) AND (NOT "ROLL_State".M[53, 6]) AND "ROLL_State".M[31, 5] AND "ROLL_State".M[35, 2] AND "ROLL_State".M[37, 0]);
   IF #r THEN
       "ROLL_State".M[37, 1] := TRUE;
   END_IF;
   #r := ("ROLL_State".M[32, 2] OR "ROLL_State".M[37, 2] OR "ROLL_State".M[39, 6]);
   IF #r THEN
       "ROLL_State".M[37, 1] := FALSE;
   END_IF;
   // PB9, STEP 5 network 8
   #r := ((NOT "ROLL_IO".Output[113, 3]) AND (NOT "ROLL_State".M[9, 1]) AND (("ROLL_IO".Input[0, 5] AND "ROLL_IO".Input[14, 3] AND "ROLL_State".M[0, 4]) OR ("ROLL_IO".Input[123, 4] AND "ROLL_IO".Input[124, 4] AND "ROLL_State".M[0, 3])) AND "ROLL_State".M[35, 2] AND "ROLL_State".M[37, 1]);
   IF #r THEN
       "ROLL_State".M[37, 2] := TRUE;
   END_IF;
   #r := ("ROLL_State".M[32, 2] OR "ROLL_State".M[37, 3]);
   IF #r THEN
       "ROLL_State".M[37, 2] := FALSE;
   END_IF;
   // PB9, STEP 5 network 9
   #r := ((NOT "ROLL_State".M[16, 0]) AND (NOT "ROLL_State".M[16, 1]) AND (NOT "ROLL_State".M[16, 4]) AND (NOT "ROLL_State".M[191, 5]) AND "ROLL_IO".Input[14, 0] AND "ROLL_State".M[190, 1] AND "ROLL_State".M[191, 4] AND "ROLL_State".M[35, 2] AND "ROLL_State".M[37, 2]);
   IF #r THEN
       "ROLL_State".M[37, 3] := TRUE;
   END_IF;
   #r := ("ROLL_State".M[32, 2] OR "ROLL_State".M[37, 5] OR "ROLL_State".M[40, 0]);
   IF #r THEN
       "ROLL_State".M[37, 3] := FALSE;
   END_IF;
   // PB9, STEP 5 network 10
   #r := ((NOT "ROLL_IO".Input[123, 5]) AND (NOT "ROLL_IO".Input[123, 6]) AND "ROLL_IO".Input[124, 1] AND "ROLL_IO".Input[124, 4] AND "ROLL_State".M[0, 3] AND "ROLL_State".M[35, 2] AND "ROLL_State".M[37, 3]);
   IF #r THEN
       "ROLL_State".M[37, 5] := TRUE;
   END_IF;
   #r := ("ROLL_State".M[32, 2] OR "ROLL_State".M[37, 6]);
   IF #r THEN
       "ROLL_State".M[37, 5] := FALSE;
   END_IF;
   // PB9, STEP 5 network 11
   #r := ((NOT "ROLL_IO".Output[113, 2]) AND "ROLL_IO".Output[113, 3] AND "ROLL_State".M[35, 2] AND "ROLL_State".M[37, 5] AND "ROLL_State".S5Timers[18].Q);
   IF #r THEN
       "ROLL_State".M[37, 6] := TRUE;
   END_IF;
   #r := ("ROLL_State".M[32, 2] OR "ROLL_State".M[37, 7]);
   IF #r THEN
       "ROLL_State".M[37, 6] := FALSE;
   END_IF;
   // PB9, STEP 5 network 12
   #r := ((NOT "ROLL_State".M[37, 5]) AND "ROLL_State".M[35, 2] AND "ROLL_State".M[37, 6]);
   IF #r THEN
       "ROLL_State".M[37, 7] := TRUE;
   END_IF;
   #r := ("ROLL_State".M[32, 2] OR "ROLL_State".M[38, 0]);
   IF #r THEN
       "ROLL_State".M[37, 7] := FALSE;
   END_IF;
   // PB9, STEP 5 network 13
   #r := ((NOT "ROLL_State".M[70, 2]) AND (((NOT "ROLL_IO".Output[113, 2]) AND "ROLL_IO".Output[113, 3] AND "ROLL_IO".Input[124, 4] AND "ROLL_State".M[28, 4] AND "ROLL_State".M[37, 0]) OR ("ROLL_State".M[37, 7] AND "ROLL_State".S5Timers[20].Q)) AND "ROLL_IO".Input[123, 5] AND "ROLL_State".M[35, 2]);
   IF #r THEN
       "ROLL_State".M[38, 0] := TRUE;
   END_IF;
   #r := ("ROLL_State".M[32, 2] OR "ROLL_State".M[39, 4]);
   IF #r THEN
       "ROLL_State".M[38, 0] := FALSE;
   END_IF;
   // PB9, STEP 5 network 14
   #r := ((NOT "ROLL_IO".Input[124, 5]) AND "ROLL_IO".Input[124, 4] AND "ROLL_State".M[35, 2] AND "ROLL_State".M[38, 0]);
   IF #r THEN
       "ROLL_State".M[39, 4] := TRUE;
   END_IF;
   #r := ("ROLL_State".M[32, 2] OR "ROLL_State".M[39, 5]);
   IF #r THEN
       "ROLL_State".M[39, 4] := FALSE;
   END_IF;
   // PB9, STEP 5 network 15
   #r := ((NOT "ROLL_IO".Input[124, 4]) AND (("ROLL_State".M[28, 4] AND "ROLL_State".M[37, 0]) OR "ROLL_State".M[39, 4]) AND "ROLL_IO".Input[124, 5] AND "ROLL_State".M[35, 2]);
   IF #r THEN
       "ROLL_State".M[39, 5] := TRUE;
   END_IF;
   #r := ("ROLL_State".M[32, 2] OR "ROLL_State".M[39, 6]);
   IF #r THEN
       "ROLL_State".M[39, 5] := FALSE;
   END_IF;
   // PB9, STEP 5 network 16
   #r := ((NOT "ROLL_IO".Input[124, 2]) AND "ROLL_IO".Input[11, 0] AND "ROLL_IO".Input[11, 6] AND "ROLL_IO".Input[12, 1] AND "ROLL_IO".Input[12, 7] AND "ROLL_IO".Input[124, 1] AND "ROLL_State".M[35, 2] AND "ROLL_State".M[39, 5]);
   IF #r THEN
       "ROLL_State".M[39, 6] := TRUE;
   END_IF;
   #r := ("ROLL_State".M[32, 2] OR "ROLL_State".M[39, 7]);
   IF #r THEN
       "ROLL_State".M[39, 6] := FALSE;
   END_IF;
   // PB9, STEP 5 network 17
   #r := ((NOT "ROLL_IO".Input[124, 1]) AND "ROLL_IO".Input[124, 2] AND "ROLL_State".M[35, 2] AND "ROLL_State".M[39, 6]);
   IF #r THEN
       "ROLL_State".M[39, 7] := TRUE;
   END_IF;
   #r := ("ROLL_State".M[32, 2] OR "ROLL_State".M[40, 0]);
   IF #r THEN
       "ROLL_State".M[39, 7] := FALSE;
   END_IF;
   // PB9, STEP 5 network 18
   #r := ((NOT "ROLL_IO".Input[12, 5]) AND ("ROLL_State".M[37, 3] OR "ROLL_State".M[39, 7]) AND "ROLL_IO".Input[11, 0] AND "ROLL_IO".Input[11, 6] AND "ROLL_IO".Input[12, 1] AND "ROLL_IO".Input[12, 7] AND "ROLL_State".M[35, 2]);
   IF #r THEN
       "ROLL_State".M[40, 0] := TRUE;
   END_IF;
   #r := ("ROLL_State".M[32, 2] OR "ROLL_State".M[40, 1]);
   IF #r THEN
       "ROLL_State".M[40, 0] := FALSE;
   END_IF;
   // PB9, STEP 5 network 19
   #r := ("ROLL_IO".Input[12, 5] AND "ROLL_IO".Input[12, 7] AND "ROLL_State".M[35, 2] AND "ROLL_State".M[40, 0]);
   IF #r THEN
       "ROLL_State".M[40, 1] := TRUE;
   END_IF;
   #r := ("ROLL_State".M[32, 2] OR "ROLL_State".M[40, 2] OR "ROLL_State".M[41, 6] OR "ROLL_State".M[43, 2] OR "ROLL_State".M[44, 7] OR "ROLL_State".M[46, 2] OR "ROLL_State".M[47, 6] OR "ROLL_State".M[49, 2] OR "ROLL_State".M[50, 6]);
   IF #r THEN
       "ROLL_State".M[40, 1] := FALSE;
   END_IF;
   // PB9, STEP 5 network 20
   #r := ((NOT "ROLL_IO".Input[11, 1]) AND "ROLL_IO".Input[11, 0] AND "ROLL_State".M[110, 0] AND "ROLL_State".M[35, 2] AND "ROLL_State".M[40, 1] AND "ROLL_State".M[63, 1]);
   IF #r THEN
       "ROLL_State".M[40, 2] := TRUE;
   END_IF;
   #r := ("ROLL_State".M[32, 2] OR "ROLL_State".M[40, 3]);
   IF #r THEN
       "ROLL_State".M[40, 2] := FALSE;
   END_IF;
   // PB9, STEP 5 network 21
   #r := ("ROLL_IO".Input[11, 1] AND "ROLL_IO".Input[11, 6] AND "ROLL_State".M[35, 2] AND "ROLL_State".M[40, 2]);
   IF #r THEN
       "ROLL_State".M[40, 3] := TRUE;
   END_IF;
   #r := ("ROLL_State".M[32, 2] OR "ROLL_State".M[40, 4]);
   IF #r THEN
       "ROLL_State".M[40, 3] := FALSE;
   END_IF;
   // PB9, STEP 5 network 22
   #r := ((NOT "ROLL_IO".Input[12, 1]) AND "ROLL_IO".Input[12, 5] AND "ROLL_State".M[35, 2] AND "ROLL_State".M[40, 3]);
   IF #r THEN
       "ROLL_State".M[40, 4] := TRUE;
   END_IF;
   #r := ("ROLL_State".M[32, 2] OR "ROLL_State".M[40, 5]);
   IF #r THEN
       "ROLL_State".M[40, 4] := FALSE;
   END_IF;
   // PB9, STEP 5 network 23
   #r := ("ROLL_IO".Input[12, 1] AND "ROLL_IO".Input[12, 7] AND "ROLL_State".M[35, 2] AND "ROLL_State".M[40, 4]);
   IF #r THEN
       "ROLL_State".M[40, 5] := TRUE;
   END_IF;
   #r := ("ROLL_State".M[32, 2] OR "ROLL_State".M[40, 6]);
   IF #r THEN
       "ROLL_State".M[40, 5] := FALSE;
   END_IF;
   // PB9, STEP 5 network 24
   #r := ("ROLL_State".M[35, 2] AND "ROLL_State".M[40, 5] AND "ROLL_State".S5Timers[1].Q);
   IF #r THEN
       "ROLL_State".M[40, 6] := TRUE;
   END_IF;
   #r := ("ROLL_State".M[32, 2] OR "ROLL_State".M[40, 7]);
   IF #r THEN
       "ROLL_State".M[40, 6] := FALSE;
   END_IF;
   // PB9, STEP 5 network 25
   #r := ("ROLL_State".M[35, 2] AND "ROLL_State".M[40, 6]);
   IF #r THEN
       "ROLL_State".M[40, 7] := TRUE;
   END_IF;
   #r := ("ROLL_State".M[32, 2] OR "ROLL_State".M[41, 0]);
   IF #r THEN
       "ROLL_State".M[40, 7] := FALSE;
   END_IF;
   // PB9, STEP 5 network 26
   #r := ((NOT "ROLL_IO".Input[12, 5]) AND (("ROLL_IO".Input[13, 3] AND "ROLL_State".M[63, 1]) OR (NOT "ROLL_State".M[111, 5])) AND "ROLL_State".M[35, 2] AND "ROLL_State".M[40, 7]);
   IF #r THEN
       "ROLL_State".M[41, 0] := TRUE;
   END_IF;
   #r := ("ROLL_State".M[32, 2] OR "ROLL_State".M[41, 1]);
   IF #r THEN
       "ROLL_State".M[41, 0] := FALSE;
   END_IF;
   // PB9, STEP 5 network 27
   #r := ("ROLL_IO".Input[12, 5] AND "ROLL_IO".Input[12, 7] AND "ROLL_State".M[35, 2] AND "ROLL_State".M[41, 0]);
   IF #r THEN
       "ROLL_State".M[41, 1] := TRUE;
   END_IF;
   #r := ("ROLL_State".M[32, 2] OR "ROLL_State".M[41, 2]);
   IF #r THEN
       "ROLL_State".M[41, 1] := FALSE;
   END_IF;
   // PB9, STEP 5 network 28
   #r := ("ROLL_State".M[35, 2] AND "ROLL_State".M[41, 1] AND "ROLL_State".S5Timers[2].Q);
   IF #r THEN
       "ROLL_State".M[41, 2] := TRUE;
   END_IF;
   #r := ("ROLL_State".M[32, 2] OR "ROLL_State".M[41, 3] OR "ROLL_State".M[41, 6] OR "ROLL_State".M[43, 2] OR "ROLL_State".M[44, 7] OR "ROLL_State".M[46, 2] OR "ROLL_State".M[47, 6] OR "ROLL_State".M[49, 2]);
   IF #r THEN
       "ROLL_State".M[41, 2] := FALSE;
   END_IF;
   // PB9, STEP 5 network 29
   #r := ((NOT "ROLL_State".M[110, 1]) AND (NOT "ROLL_State".M[110, 2]) AND "ROLL_State".M[35, 2] AND "ROLL_State".M[41, 2]);
   IF #r THEN
       "ROLL_State".M[41, 3] := TRUE;
   END_IF;
   #r := ("ROLL_State".M[32, 2] OR "ROLL_State".M[41, 4]);
   IF #r THEN
       "ROLL_State".M[41, 3] := FALSE;
   END_IF;
   // PB9, STEP 5 network 30
   #r := ("ROLL_IO".Input[13, 3] AND "ROLL_State".M[35, 2] AND "ROLL_State".M[41, 3] AND "ROLL_State".M[63, 1]);
   IF #r THEN
       "ROLL_State".M[41, 4] := TRUE;
   END_IF;
   #r := ("ROLL_State".M[32, 2] OR "ROLL_State".M[44, 7] OR "ROLL_State".M[50, 6] OR "ROLL_State".M[52, 0]);
   IF #r THEN
       "ROLL_State".M[41, 4] := FALSE;
   END_IF;
   // PB9, STEP 5 network 31
   #r := ((NOT "ROLL_IO".Input[11, 2]) AND (((NOT "ROLL_State".M[110, 0]) AND "ROLL_State".M[40, 1]) OR "ROLL_State".M[41, 2]) AND "ROLL_IO".Input[12, 5] AND "ROLL_IO".Input[12, 7] AND "ROLL_State".M[110, 1] AND "ROLL_State".M[35, 2]);
   IF #r THEN
       "ROLL_State".M[41, 6] := TRUE;
   END_IF;
   #r := ("ROLL_State".M[32, 2] OR "ROLL_State".M[41, 7]);
   IF #r THEN
       "ROLL_State".M[41, 6] := FALSE;
   END_IF;
   // PB9, STEP 5 network 32
   #r := ("ROLL_IO".Input[11, 2] AND "ROLL_IO".Input[11, 6] AND "ROLL_State".M[35, 2] AND "ROLL_State".M[41, 6]);
   IF #r THEN
       "ROLL_State".M[41, 7] := TRUE;
   END_IF;
   #r := ("ROLL_State".M[32, 2] OR "ROLL_State".M[42, 0]);
   IF #r THEN
       "ROLL_State".M[41, 7] := FALSE;
   END_IF;
   // PB9, STEP 5 network 33
   #r := ((NOT "ROLL_IO".Input[12, 1]) AND "ROLL_IO".Input[12, 5] AND "ROLL_State".M[35, 2] AND "ROLL_State".M[41, 7]);
   IF #r THEN
       "ROLL_State".M[42, 0] := TRUE;
   END_IF;
   #r := ("ROLL_State".M[32, 2] OR "ROLL_State".M[42, 1]);
   IF #r THEN
       "ROLL_State".M[42, 0] := FALSE;
   END_IF;
   // PB9, STEP 5 network 34
   #r := ("ROLL_IO".Input[12, 1] AND "ROLL_IO".Input[12, 7] AND "ROLL_State".M[35, 2] AND "ROLL_State".M[42, 0]);
   IF #r THEN
       "ROLL_State".M[42, 1] := TRUE;
   END_IF;
   #r := ("ROLL_State".M[32, 2] OR "ROLL_State".M[42, 2]);
   IF #r THEN
       "ROLL_State".M[42, 1] := FALSE;
   END_IF;
   // PB9, STEP 5 network 35
   #r := ("ROLL_State".M[35, 2] AND "ROLL_State".M[42, 1] AND "ROLL_State".S5Timers[1].Q);
   IF #r THEN
       "ROLL_State".M[42, 2] := TRUE;
   END_IF;
   #r := ("ROLL_State".M[32, 2] OR "ROLL_State".M[42, 3]);
   IF #r THEN
       "ROLL_State".M[42, 2] := FALSE;
   END_IF;
   // PB9, STEP 5 network 36
   #r := ("ROLL_State".M[35, 2] AND "ROLL_State".M[42, 2]);
   IF #r THEN
       "ROLL_State".M[42, 3] := TRUE;
   END_IF;
   #r := ("ROLL_State".M[32, 2] OR "ROLL_State".M[42, 4]);
   IF #r THEN
       "ROLL_State".M[42, 3] := FALSE;
   END_IF;
   // PB9, STEP 5 network 37
   #r := ((NOT "ROLL_IO".Input[12, 5]) AND (("ROLL_IO".Input[13, 3] AND "ROLL_State".M[63, 1]) OR (NOT "ROLL_State".M[111, 5])) AND "ROLL_State".M[35, 2] AND "ROLL_State".M[42, 3]);
   IF #r THEN
       "ROLL_State".M[42, 4] := TRUE;
   END_IF;
   #r := ("ROLL_State".M[32, 2] OR "ROLL_State".M[42, 5]);
   IF #r THEN
       "ROLL_State".M[42, 4] := FALSE;
   END_IF;
   // PB9, STEP 5 network 38
   #r := ("ROLL_IO".Input[12, 5] AND "ROLL_IO".Input[12, 7] AND "ROLL_State".M[35, 2] AND "ROLL_State".M[42, 4]);
   IF #r THEN
       "ROLL_State".M[42, 5] := TRUE;
   END_IF;
   #r := ("ROLL_State".M[32, 2] OR "ROLL_State".M[42, 6]);
   IF #r THEN
       "ROLL_State".M[42, 5] := FALSE;
   END_IF;
   // PB9, STEP 5 network 39
   #r := ("ROLL_State".M[35, 2] AND "ROLL_State".M[42, 5] AND "ROLL_State".S5Timers[2].Q);
   IF #r THEN
       "ROLL_State".M[42, 6] := TRUE;
   END_IF;
   #r := ("ROLL_State".M[32, 2] OR "ROLL_State".M[42, 7] OR "ROLL_State".M[43, 2] OR "ROLL_State".M[44, 7] OR "ROLL_State".M[46, 2] OR "ROLL_State".M[47, 6] OR "ROLL_State".M[49, 2]);
   IF #r THEN
       "ROLL_State".M[42, 6] := FALSE;
   END_IF;
   // PB9, STEP 5 network 40
   #r := ((NOT "ROLL_State".M[110, 2]) AND "ROLL_State".M[35, 2] AND "ROLL_State".M[42, 6]);
   IF #r THEN
       "ROLL_State".M[42, 7] := TRUE;
   END_IF;
   #r := ("ROLL_State".M[32, 2] OR "ROLL_State".M[43, 0]);
   IF #r THEN
       "ROLL_State".M[42, 7] := FALSE;
   END_IF;
   // PB9, STEP 5 network 41
   #r := ("ROLL_IO".Input[13, 3] AND "ROLL_State".M[35, 2] AND "ROLL_State".M[42, 7] AND "ROLL_State".M[63, 1]);
   IF #r THEN
       "ROLL_State".M[43, 0] := TRUE;
   END_IF;
   #r := ("ROLL_State".M[32, 2] OR "ROLL_State".M[44, 7] OR "ROLL_State".M[50, 6] OR "ROLL_State".M[52, 0]);
   IF #r THEN
       "ROLL_State".M[43, 0] := FALSE;
   END_IF;
   // PB9, STEP 5 network 42
   #r := ((NOT "ROLL_IO".Input[11, 3]) AND (((NOT "ROLL_State".M[110, 0]) AND (NOT "ROLL_State".M[110, 1]) AND "ROLL_State".M[40, 1]) OR ((NOT "ROLL_State".M[110, 1]) AND "ROLL_State".M[41, 2]) OR "ROLL_State".M[42, 6]) AND "ROLL_IO".Input[12, 5] AND "ROLL_IO".Input[12, 7] AND "ROLL_State".M[110, 2] AND "ROLL_State".M[35, 2]);
   IF #r THEN
       "ROLL_State".M[43, 2] := TRUE;
   END_IF;
   #r := ("ROLL_State".M[32, 2] OR "ROLL_State".M[43, 3]);
   IF #r THEN
       "ROLL_State".M[43, 2] := FALSE;
   END_IF;
   // PB9, STEP 5 network 43
   #r := ("ROLL_IO".Input[11, 3] AND "ROLL_IO".Input[11, 6] AND "ROLL_State".M[35, 2] AND "ROLL_State".M[43, 2]);
   IF #r THEN
       "ROLL_State".M[43, 3] := TRUE;
   END_IF;
   #r := ("ROLL_State".M[32, 2] OR "ROLL_State".M[43, 4]);
   IF #r THEN
       "ROLL_State".M[43, 3] := FALSE;
   END_IF;
   // PB9, STEP 5 network 44
   #r := ((NOT "ROLL_IO".Input[12, 1]) AND "ROLL_IO".Input[12, 5] AND "ROLL_State".M[35, 2] AND "ROLL_State".M[43, 3]);
   IF #r THEN
       "ROLL_State".M[43, 4] := TRUE;
   END_IF;
   #r := ("ROLL_State".M[32, 2] OR "ROLL_State".M[43, 5]);
   IF #r THEN
       "ROLL_State".M[43, 4] := FALSE;
   END_IF;
   // PB9, STEP 5 network 45
   #r := ("ROLL_IO".Input[12, 1] AND "ROLL_IO".Input[12, 7] AND "ROLL_State".M[35, 2] AND "ROLL_State".M[43, 4]);
   IF #r THEN
       "ROLL_State".M[43, 5] := TRUE;
   END_IF;
   #r := ("ROLL_State".M[32, 2] OR "ROLL_State".M[43, 6]);
   IF #r THEN
       "ROLL_State".M[43, 5] := FALSE;
   END_IF;
   // PB9, STEP 5 network 46
   #r := ("ROLL_State".M[35, 2] AND "ROLL_State".M[43, 5] AND "ROLL_State".S5Timers[1].Q);
   IF #r THEN
       "ROLL_State".M[43, 6] := TRUE;
   END_IF;
   #r := ("ROLL_State".M[32, 2] OR "ROLL_State".M[43, 7]);
   IF #r THEN
       "ROLL_State".M[43, 6] := FALSE;
   END_IF;
   // PB9, STEP 5 network 47
   #r := ("ROLL_State".M[35, 2] AND "ROLL_State".M[43, 6]);
   IF #r THEN
       "ROLL_State".M[43, 7] := TRUE;
   END_IF;
   #r := ("ROLL_State".M[32, 2] OR "ROLL_State".M[44, 0]);
   IF #r THEN
       "ROLL_State".M[43, 7] := FALSE;
   END_IF;
   // PB9, STEP 5 network 48
   #r := ((NOT "ROLL_IO".Input[12, 5]) AND (("ROLL_IO".Input[13, 3] AND "ROLL_State".M[63, 1]) OR (NOT "ROLL_State".M[111, 5])) AND "ROLL_State".M[35, 2] AND "ROLL_State".M[43, 7]);
   IF #r THEN
       "ROLL_State".M[44, 0] := TRUE;
   END_IF;
   #r := ("ROLL_State".M[32, 2] OR "ROLL_State".M[44, 1]);
   IF #r THEN
       "ROLL_State".M[44, 0] := FALSE;
   END_IF;
   // PB9, STEP 5 network 49
   #r := ("ROLL_IO".Input[12, 5] AND "ROLL_IO".Input[12, 7] AND "ROLL_State".M[35, 2] AND "ROLL_State".M[44, 0]);
   IF #r THEN
       "ROLL_State".M[44, 1] := TRUE;
   END_IF;
   #r := ("ROLL_State".M[32, 2] OR "ROLL_State".M[44, 2]);
   IF #r THEN
       "ROLL_State".M[44, 1] := FALSE;
   END_IF;
   // PB9, STEP 5 network 50
   #r := ("ROLL_State".M[35, 2] AND "ROLL_State".M[44, 1] AND "ROLL_State".S5Timers[2].Q);
   IF #r THEN
       "ROLL_State".M[44, 2] := TRUE;
   END_IF;
   #r := ("ROLL_State".M[32, 2] OR "ROLL_State".M[44, 3] OR "ROLL_State".M[44, 7] OR "ROLL_State".M[46, 2] OR "ROLL_State".M[47, 6] OR "ROLL_State".M[49, 2]);
   IF #r THEN
       "ROLL_State".M[44, 2] := FALSE;
   END_IF;
   // PB9, STEP 5 network 51
   #r := ("ROLL_State".M[35, 2] AND "ROLL_State".M[44, 2]);
   IF #r THEN
       "ROLL_State".M[44, 3] := TRUE;
   END_IF;
   #r := ("ROLL_State".M[32, 2] OR "ROLL_State".M[44, 4]);
   IF #r THEN
       "ROLL_State".M[44, 3] := FALSE;
   END_IF;
   // PB9, STEP 5 network 52
   #r := ("ROLL_IO".Input[13, 3] AND "ROLL_State".M[35, 2] AND "ROLL_State".M[44, 3] AND "ROLL_State".M[63, 1]);
   IF #r THEN
       "ROLL_State".M[44, 4] := TRUE;
   END_IF;
   #r := ("ROLL_State".M[32, 2] OR "ROLL_State".M[44, 7] OR "ROLL_State".M[50, 6] OR "ROLL_State".M[52, 0]);
   IF #r THEN
       "ROLL_State".M[44, 4] := FALSE;
   END_IF;
   // PB9, STEP 5 network 53
   #r := (((NOT "ROLL_State".M[110, 0]) AND (NOT "ROLL_State".M[110, 1]) AND (NOT "ROLL_State".M[110, 2]) AND "ROLL_State".M[40, 1]) OR ((NOT "ROLL_State".M[110, 1]) AND (NOT "ROLL_State".M[110, 2]) AND "ROLL_State".M[41, 4]) OR ((NOT "ROLL_State".M[110, 2]) AND "ROLL_State".M[43, 0]) OR "ROLL_State".M[44, 4]);
   "ROLL_State".M[240, 0] := #r;
   // PB9, STEP 5 network 54
   #r := ((NOT "ROLL_IO".Input[11, 4]) AND "ROLL_IO".Input[12, 5] AND "ROLL_IO".Input[12, 7] AND "ROLL_State".M[110, 3] AND "ROLL_State".M[240, 0] AND "ROLL_State".M[35, 2] AND "ROLL_State".M[63, 1]);
   IF #r THEN
       "ROLL_State".M[44, 7] := TRUE;
   END_IF;
   #r := ("ROLL_State".M[32, 2] OR "ROLL_State".M[45, 0]);
   IF #r THEN
       "ROLL_State".M[44, 7] := FALSE;
   END_IF;
   // PB9, STEP 5 network 55
   #r := ("ROLL_IO".Input[11, 4] AND "ROLL_IO".Input[11, 6] AND "ROLL_State".M[35, 2] AND "ROLL_State".M[44, 7]);
   IF #r THEN
       "ROLL_State".M[45, 0] := TRUE;
   END_IF;
   #r := ("ROLL_State".M[32, 2] OR "ROLL_State".M[45, 1]);
   IF #r THEN
       "ROLL_State".M[45, 0] := FALSE;
   END_IF;
   // PB9, STEP 5 network 56
   #r := ((NOT "ROLL_IO".Input[12, 1]) AND "ROLL_IO".Input[12, 5] AND "ROLL_State".M[35, 2] AND "ROLL_State".M[45, 0]);
   IF #r THEN
       "ROLL_State".M[45, 1] := TRUE;
   END_IF;
   #r := ("ROLL_State".M[32, 2] OR "ROLL_State".M[45, 2]);
   IF #r THEN
       "ROLL_State".M[45, 1] := FALSE;
   END_IF;
   // PB9, STEP 5 network 57
   #r := ("ROLL_IO".Input[12, 1] AND "ROLL_IO".Input[12, 7] AND "ROLL_State".M[35, 2] AND "ROLL_State".M[45, 1]);
   IF #r THEN
       "ROLL_State".M[45, 2] := TRUE;
   END_IF;
   #r := ("ROLL_State".M[32, 2] OR "ROLL_State".M[45, 3]);
   IF #r THEN
       "ROLL_State".M[45, 2] := FALSE;
   END_IF;
   // PB9, STEP 5 network 58
   #r := ("ROLL_State".M[35, 2] AND "ROLL_State".M[45, 2] AND "ROLL_State".S5Timers[1].Q);
   IF #r THEN
       "ROLL_State".M[45, 3] := TRUE;
   END_IF;
   #r := ("ROLL_State".M[32, 2] OR "ROLL_State".M[45, 4]);
   IF #r THEN
       "ROLL_State".M[45, 3] := FALSE;
   END_IF;
   // PB9, STEP 5 network 59
   #r := ("ROLL_State".M[35, 2] AND "ROLL_State".M[45, 3]);
   IF #r THEN
       "ROLL_State".M[45, 4] := TRUE;
   END_IF;
   #r := ("ROLL_State".M[32, 2] OR "ROLL_State".M[45, 5]);
   IF #r THEN
       "ROLL_State".M[45, 4] := FALSE;
   END_IF;
   // PB9, STEP 5 network 60
   #r := ((NOT "ROLL_IO".Input[12, 5]) AND "ROLL_State".M[35, 2] AND "ROLL_State".M[45, 4]);
   IF #r THEN
       "ROLL_State".M[45, 5] := TRUE;
   END_IF;
   #r := ("ROLL_State".M[32, 2] OR "ROLL_State".M[45, 6]);
   IF #r THEN
       "ROLL_State".M[45, 5] := FALSE;
   END_IF;
   // PB9, STEP 5 network 61
   #r := ("ROLL_IO".Input[12, 5] AND "ROLL_IO".Input[12, 7] AND "ROLL_State".M[35, 2] AND "ROLL_State".M[45, 5]);
   IF #r THEN
       "ROLL_State".M[45, 6] := TRUE;
   END_IF;
   #r := ("ROLL_State".M[32, 2] OR "ROLL_State".M[45, 7]);
   IF #r THEN
       "ROLL_State".M[45, 6] := FALSE;
   END_IF;
   // PB9, STEP 5 network 62
   #r := (("ROLL_State".M[0, 4] OR "ROLL_State".S5Timers[2].Q) AND "ROLL_State".M[35, 2] AND "ROLL_State".M[45, 6]);
   IF #r THEN
       "ROLL_State".M[45, 7] := TRUE;
   END_IF;
   #r := ("ROLL_State".M[32, 2] OR "ROLL_State".M[46, 0] OR "ROLL_State".M[46, 2] OR "ROLL_State".M[47, 6] OR "ROLL_State".M[49, 2]);
   IF #r THEN
       "ROLL_State".M[45, 7] := FALSE;
   END_IF;
   // PB9, STEP 5 network 63
   #r := ("ROLL_State".M[35, 2] AND "ROLL_State".M[45, 7]);
   IF #r THEN
       "ROLL_State".M[46, 0] := TRUE;
   END_IF;
   #r := ("ROLL_State".M[32, 2] OR "ROLL_State".M[46, 1]);
   IF #r THEN
       "ROLL_State".M[46, 0] := FALSE;
   END_IF;
   // PB9, STEP 5 network 64
   #r := ("ROLL_IO".Input[13, 3] AND "ROLL_State".M[35, 2] AND "ROLL_State".M[46, 0] AND "ROLL_State".M[63, 1]);
   IF #r THEN
       "ROLL_State".M[46, 1] := TRUE;
   END_IF;
   #r := ("ROLL_State".M[32, 2] OR "ROLL_State".M[50, 6] OR "ROLL_State".M[52, 0]);
   IF #r THEN
       "ROLL_State".M[46, 1] := FALSE;
   END_IF;
   // PB9, STEP 5 network 65
   RETURN;
END_FUNCTION

FUNCTION "ROLL_ReadInputs" : Void   // FC36, SCL
{ S7_Optimized_Access := 'TRUE' }
VERSION : 0.1
// stored: AutoNumber true, IsIECCheckEnabled false, SetENOAutomatically false, UDAEnableTagReadback false
   VAR_TEMP
      "b" : Int;
      bit : Int;
   END_VAR
BEGIN

   // Confirmed four-station profile: absent optional inputs are zero.
   FOR #b := 119 TO 125 DO
       FOR #bit := 0 TO 7 DO
           "ROLL_IO".Input[#b, #bit] := FALSE;
       END_FOR;
   END_FOR;
   IF "ROLL_IO".PhysicalIoConfigured AND NOT "ROLL_IO".Simulation THEN
       "ROLL_IO".Input[0, 0] := "Tag__639276557951123186";
       "ROLL_IO".Input[0, 1] := "Tag__639276557952818668";
       "ROLL_IO".Input[0, 2] := "Tag__639276557952918398";
       "ROLL_IO".Input[0, 3] := "Tag__639276557952998183";
       "ROLL_IO".Input[0, 4] := "Tag__639276557953077986";
       "ROLL_IO".Input[0, 5] := "Tag__639276557953157762";
       "ROLL_IO".Input[0, 6] := "Tag__639276557953227573";
       "ROLL_IO".Input[0, 7] := "Tag__639276557953307358";
       "ROLL_IO".Input[1, 0] := "Tag__639276557953367206";
       "ROLL_IO".Input[1, 1] := "Tag__639276557953447409";
       "ROLL_IO".Input[1, 2] := "Tag__639276557953526828";
       "ROLL_IO".Input[1, 3] := "Tag__639276557953606562";
       "ROLL_IO".Input[1, 4] := "Tag__639276557953686353";
       "ROLL_IO".Input[1, 5] := "Tag__639276557953766129";
       "ROLL_IO".Input[1, 6] := "Tag__639276557953835956";
       "ROLL_IO".Input[1, 7] := "Tag__639276557953915729";
       "ROLL_IO".Input[2, 0] := "Tag__639276557953985541";
       "ROLL_IO".Input[2, 1] := "Tag__639276557954055362";
       "ROLL_IO".Input[2, 2] := "Tag__639276557954135145";
       "ROLL_IO".Input[2, 3] := "Tag__639276557954204958";
       "ROLL_IO".Input[2, 4] := "Tag__639276557954284740";
       "ROLL_IO".Input[2, 5] := "Tag__639276557954354781";
       "ROLL_IO".Input[2, 6] := "Tag__639276557954434344";
       "ROLL_IO".Input[2, 7] := "Tag__639276557954494175";
       "ROLL_IO".Input[3, 0] := "Tag__639276557954554015";
       "ROLL_IO".Input[3, 1] := "Tag__639276557954604247";
       "ROLL_IO".Input[3, 2] := "Tag__639276557954663730";
       "ROLL_IO".Input[3, 3] := "Tag__639276557954723560";
       "ROLL_IO".Input[3, 4] := "Tag__639276557954773427";
       "ROLL_IO".Input[3, 5] := "Tag__639276557954833268";
       "ROLL_IO".Input[3, 6] := "Tag__639276557954893102";
       "ROLL_IO".Input[3, 7] := "Tag__639276557954953006";
       "ROLL_IO".Input[4, 0] := "Tag__639276557955012796";
       "ROLL_IO".Input[4, 1] := "Tag__639276557955062653";
       "ROLL_IO".Input[4, 2] := "Tag__639276557955122494";
       "ROLL_IO".Input[4, 3] := "Tag__639276557955182529";
       "ROLL_IO".Input[4, 4] := "Tag__639276557955242183";
       "ROLL_IO".Input[4, 5] := "Tag__639276557955302013";
       "ROLL_IO".Input[4, 6] := "Tag__639276557955362031";
       "ROLL_IO".Input[4, 7] := "Tag__639276557955411719";
       "ROLL_IO".Input[5, 0] := "Tag__639276557955481879";
       "ROLL_IO".Input[5, 1] := "Tag__639276557955541374";
       "ROLL_IO".Input[5, 2] := "Tag__639276557955601431";
       "ROLL_IO".Input[5, 3] := "Tag__639276557955661053";
       "ROLL_IO".Input[5, 4] := "Tag__639276557955710919";
       "ROLL_IO".Input[5, 5] := "Tag__639276557955770760";
       "ROLL_IO".Input[5, 6] := "Tag__639276557955820633";
       "ROLL_IO".Input[5, 7] := "Tag__639276557955880472";
       "ROLL_IO".Input[6, 0] := "Tag__639276557955940421";
       "ROLL_IO".Input[6, 1] := "Tag__639276557955990183";
       "ROLL_IO".Input[6, 2] := "Tag__639276557956050021";
       "ROLL_IO".Input[6, 3] := "Tag__639276557956099878";
       "ROLL_IO".Input[6, 4] := "Tag__639276557956149744";
       "ROLL_IO".Input[6, 5] := "Tag__639276557956209908";
       "ROLL_IO".Input[6, 6] := "Tag__639276557956259702";
       "ROLL_IO".Input[6, 7] := "Tag__639276557956319298";
       "ROLL_IO".Input[7, 0] := "Tag__639276557956369159";
       "ROLL_IO".Input[7, 1] := "Tag__639276557956419023";
       "ROLL_IO".Input[7, 2] := "Tag__639276557956479295";
       "ROLL_IO".Input[7, 3] := "Tag__639276557956528731";
       "ROLL_IO".Input[7, 4] := "Tag__639276557956578596";
       "ROLL_IO".Input[7, 5] := "Tag__639276557956638440";
       "ROLL_IO".Input[7, 6] := "Tag__639276557956698277";
       "ROLL_IO".Input[7, 7] := "Tag__639276557956758124";
       "ROLL_IO".Input[8, 0] := "Tag__639276557956808017";
       "ROLL_IO".Input[8, 1] := "Tag__639276557956867823";
       "ROLL_IO".Input[8, 2] := "Tag__639276557956917689";
       "ROLL_IO".Input[8, 3] := "Tag__639276557956977678";
       "ROLL_IO".Input[8, 4] := "Tag__639276557957037371";
       "ROLL_IO".Input[8, 5] := "Tag__639276557957087293";
       "ROLL_IO".Input[8, 6] := "Tag__639276557957147084";
       "ROLL_IO".Input[8, 7] := "Tag__639276557957196942";
       "ROLL_IO".Input[9, 0] := "Tag__639276557957256782";
       "ROLL_IO".Input[9, 1] := "Tag__639276557957316622";
       "ROLL_IO".Input[9, 2] := "Tag__639276557957366490";
       "ROLL_IO".Input[9, 3] := "Tag__639276557957426337";
       "ROLL_IO".Input[9, 4] := "Tag__639276557957476206";
       "ROLL_IO".Input[9, 5] := "Tag__639276557957526061";
       "ROLL_IO".Input[9, 6] := "Tag__639276557957586243";
       "ROLL_IO".Input[9, 7] := "Tag__639276557957645746";
       "ROLL_IO".Input[10, 0] := "Tag__639276557957705582";
       "ROLL_IO".Input[10, 1] := "Tag__639276557957755449";
       "ROLL_IO".Input[10, 2] := "Tag__639276557957805314";
       "ROLL_IO".Input[10, 3] := "Tag__639276557957865154";
       "ROLL_IO".Input[10, 4] := "Tag__639276557957915021";
       "ROLL_IO".Input[10, 5] := "Tag__639276557957964888";
       "ROLL_IO".Input[10, 6] := "Tag__639276557958024728";
       "ROLL_IO".Input[10, 7] := "Tag__639276557958074957";
       "ROLL_IO".Input[11, 0] := "Tag__639276557958124460";
       "ROLL_IO".Input[11, 1] := "Tag__639276557958184301";
       "ROLL_IO".Input[11, 2] := "Tag__639276557958234167";
       "ROLL_IO".Input[11, 3] := "Tag__639276557958294016";
       "ROLL_IO".Input[11, 4] := "Tag__639276557958343874";
       "ROLL_IO".Input[11, 5] := "Tag__639276557958393749";
       "ROLL_IO".Input[11, 6] := "Tag__639276557958453636";
       "ROLL_IO".Input[11, 7] := "Tag__639276557958503448";
       "ROLL_IO".Input[12, 0] := "Tag__639276557958553313";
       "ROLL_IO".Input[12, 1] := "Tag__639276557958613155";
       "ROLL_IO".Input[12, 2] := "Tag__639276557958663020";
       "ROLL_IO".Input[12, 3] := "Tag__639276557958712886";
       "ROLL_IO".Input[12, 4] := "Tag__639276557958772727";
       "ROLL_IO".Input[12, 5] := "Tag__639276557958822593";
       "ROLL_IO".Input[12, 6] := "Tag__639276557958902547";
       "ROLL_IO".Input[12, 7] := "Tag__639276557958962223";
       "ROLL_IO".Input[13, 0] := "Tag__639276557959022060";
       "ROLL_IO".Input[13, 1] := "Tag__639276557959071925";
       "ROLL_IO".Input[13, 2] := "Tag__639276557959131766";
       "ROLL_IO".Input[13, 3] := "Tag__639276557959191606";
       "ROLL_IO".Input[13, 4] := "Tag__639276557959251774";
       "ROLL_IO".Input[13, 5] := "Tag__639276557959311297";
       "ROLL_IO".Input[13, 6] := "Tag__639276557959371125";
       "ROLL_IO".Input[13, 7] := "Tag__639276557959430966";
       "ROLL_IO".Input[14, 0] := "Tag__639276557959490814";
       "ROLL_IO".Input[14, 1] := "Tag__639276557959540672";
       "ROLL_IO".Input[14, 2] := "Tag__639276557959600839";
       "ROLL_IO".Input[14, 3] := "Tag__639276557959650385";
       "ROLL_IO".Input[14, 4] := "Tag__639276557959710219";
       "ROLL_IO".Input[14, 5] := "Tag__639276557959760095";
       "ROLL_IO".Input[14, 6] := "Tag__639276557959809951";
       "ROLL_IO".Input[14, 7] := "Tag__639276557959869792";
       "ROLL_IO".Input[15, 0] := "Tag__639276557959929638";
       "ROLL_IO".Input[15, 1] := "Tag__639276557959979499";
       "ROLL_IO".Input[15, 2] := "Tag__639276557960039343";
       "ROLL_IO".Input[15, 3] := "Tag__639276557960089204";
       "ROLL_IO".Input[15, 4] := "Tag__639276557960139071";
       "ROLL_IO".Input[15, 5] := "Tag__639276557960198912";
       "ROLL_IO".Input[15, 6] := "Tag__639276557960248790";
       "ROLL_IO".Input[15, 7] := "Tag__639276557960308618";
   END_IF;
END_FUNCTION

FUNCTION "ROLL_SetMWord" : Void   // FC2, SCL
{ S7_Optimized_Access := 'TRUE' }
VERSION : 0.1
// stored: AutoNumber true, IsIECCheckEnabled false, SetENOAutomatically false, UDAEnableTagReadback false
   VAR_INPUT
      FirstByte : Int;
      Value : Word;
   END_VAR
   VAR_TEMP
      bit : Int;
   END_VAR
BEGIN

   IF (#FirstByte < 0) OR (#FirstByte > 254) THEN
       "ROLL_IO".ConversionFault := TRUE;
       RETURN;
   END_IF;
   FOR #bit := 0 TO 7 DO
       "ROLL_State".M[#FirstByte, #bit] := (#Value AND SHL(IN := W#16#0001, N := INT_TO_USINT(#bit + 8))) <> W#16#0000;
       "ROLL_State".M[#FirstByte + 1, #bit] := (#Value AND SHL(IN := W#16#0001, N := INT_TO_USINT(#bit))) <> W#16#0000;
   END_FOR;
END_FUNCTION

FUNCTION "ROLL_ShowRecipe" : Void   // FC11, SCL
{ S7_Optimized_Access := 'TRUE' }
VERSION : 0.1
// stored: AutoNumber true, IsIECCheckEnabled false, SetENOAutomatically false, UDAEnableTagReadback false
BEGIN

   "ROLL_HMI".CurrentProgram := "ROLL_State".CurrentProgram;
   "ROLL_HMI".SelectedProgram := "ROLL_State".CurrentProgram;
   "ROLL_HMI".Dwell1Seconds := "ROLL_DecodeBCD"(Value := "ROLL_DB205".DW[5]);
   "ROLL_HMI".Drain1Seconds := "ROLL_DecodeBCD"(Value := "ROLL_DB205".DW[9]);
   "ROLL_HMI".Dwell2Seconds := "ROLL_DecodeBCD"(Value := "ROLL_DB205".DW[17]);
   "ROLL_HMI".Drain2Seconds := "ROLL_DecodeBCD"(Value := "ROLL_DB205".DW[21]);
   "ROLL_HMI".Dwell3Seconds := "ROLL_DecodeBCD"(Value := "ROLL_DB205".DW[25]);
   "ROLL_HMI".Drain3Seconds := "ROLL_DecodeBCD"(Value := "ROLL_DB205".DW[29]);
   "ROLL_HMI".Dry4Seconds := "ROLL_DecodeBCD"(Value := "ROLL_DB205".DW[33]);
   "ROLL_HMI".Ultrasound1 := "ROLL_DB205".DW[13] = W#16#0001;
   "ROLL_HMI".BasketMotion := WORD_TO_INT("ROLL_DB205".DW[37]);
   "ROLL_HMI".BathLift := "ROLL_DB205".DW[41] = W#16#0001;
END_FUNCTION

FUNCTION "ROLL_TimerOp" : Void   // FC6, SCL
{ S7_Optimized_Access := 'TRUE' }
VERSION : 0.1
// stored: AutoNumber true, IsIECCheckEnabled false, SetENOAutomatically false, UDAEnableTagReadback false
   VAR_INPUT
      Number : Int;
      Operation : Int;   // 0=SE on-delay; 1=SA off-delay; 2=R reset
      Signal : Bool;
      Preset : Word;
   END_VAR
   VAR_TEMP
      base : Int;
      count : Int;
      trigger : Bool;
   END_VAR
BEGIN

   IF (#Number < 0) OR (#Number > 127) THEN
       "ROLL_IO".ConversionFault := TRUE;
       RETURN;
   END_IF;
   IF #Operation = 2 THEN
       IF #Signal THEN
           "ROLL_State".S5Timers[#Number].RemainingMs := 0.0;
           "ROLL_State".S5Timers[#Number].Q := FALSE;
       END_IF;
       RETURN;
   END_IF;
   #trigger := ((#Operation = 0) AND #Signal AND NOT "ROLL_State".S5Timers[#Number].Previous)
   OR ((#Operation = 1) AND NOT #Signal AND "ROLL_State".S5Timers[#Number].Previous);
   IF #trigger THEN
       #count := "ROLL_DecodeBCD"(Value := #Preset);
       #base := WORD_TO_INT(SHR(IN := #Preset AND W#16#F000, N := 12));
       CASE #base OF
           0:
               #base := 10;
           1:
               #base := 100;
           2:
               #base := 1000;
           3:
               #base := 10000;
           ELSE
               #base := 0;
       END_CASE;
       IF (#base = 0) OR (#count < 0) THEN
           "ROLL_IO".ConversionFault := TRUE;
           "ROLL_State".S5Timers[#Number].RemainingMs := 0.0;
           "ROLL_State".S5Timers[#Number].Q := FALSE;
           RETURN;
       END_IF;
       "ROLL_State".S5Timers[#Number].BaseMs := #base;
       "ROLL_State".S5Timers[#Number].RemainingMs := INT_TO_LREAL(#count) * INT_TO_LREAL(#base);
   END_IF;
   "ROLL_State".S5Timers[#Number].Mode := #Operation;
   IF #Operation = 0 THEN
       IF NOT #Signal THEN
           "ROLL_State".S5Timers[#Number].RemainingMs := 0.0;
       END_IF;
       "ROLL_State".S5Timers[#Number].Q := #Signal AND ("ROLL_State".S5Timers[#Number].RemainingMs <= 0.0);
   ELSIF #Operation = 1 THEN
       IF #Signal THEN
           "ROLL_State".S5Timers[#Number].RemainingMs := 0.0;
       END_IF;
       "ROLL_State".S5Timers[#Number].Q := #Signal OR ("ROLL_State".S5Timers[#Number].RemainingMs > 0.0);
   ELSE
       "ROLL_IO".ConversionFault := TRUE;
   END_IF;
   "ROLL_State".S5Timers[#Number].Previous := #Signal;
END_FUNCTION

FUNCTION "ROLL_TimerValue" : Word   // FC7, SCL
{ S7_Optimized_Access := 'TRUE' }
VERSION : 0.1
// stored: AutoNumber true, IsIECCheckEnabled false, SetENOAutomatically false, UDAEnableTagReadback false
   VAR_INPUT
      Number : Int;
   END_VAR
   VAR_TEMP
      count : DInt;
   END_VAR
BEGIN

   #ROLL_TimerValue := W#16#0000;
   IF (#Number < 0) OR (#Number > 127) THEN
       "ROLL_IO".ConversionFault := TRUE;
       RETURN;
   END_IF;
   IF "ROLL_State".S5Timers[#Number].BaseMs > 0 THEN
       #count := CEIL("ROLL_State".S5Timers[#Number].RemainingMs / INT_TO_LREAL("ROLL_State".S5Timers[#Number].BaseMs));
       #ROLL_TimerValue := DINT_TO_WORD(#count);
   END_IF;
END_FUNCTION

FUNCTION "ROLL_WriteOutputs" : Void   // FC37, SCL
{ S7_Optimized_Access := 'TRUE' }
VERSION : 0.1
// stored: AutoNumber true, IsIECCheckEnabled false, SetENOAutomatically false, UDAEnableTagReadback false
   VAR_TEMP
      enabled : Bool;
   END_VAR
BEGIN

   IF "ROLL_IO".PhysicalIoConfigured THEN
       #enabled := "ROLL_IO".PhysicalOutputsEnabled AND NOT "ROLL_IO".Simulation AND NOT "ROLL_IO".ConversionFault;
       "Tag__639276557961655014" := #enabled AND "ROLL_IO".Output[16, 0];
       "Tag__639276557961724830" := #enabled AND "ROLL_IO".Output[16, 1];
       "Tag__639276557961774695" := #enabled AND "ROLL_IO".Output[16, 2];
       "Tag__639276557961834550" := #enabled AND "ROLL_IO".Output[16, 3];
       "Tag__639276557961894385" := #enabled AND "ROLL_IO".Output[16, 4];
       "Tag__639276557961944242" := #enabled AND "ROLL_IO".Output[16, 5];
       "Tag__639276557962004083" := #enabled AND "ROLL_IO".Output[16, 6];
       "Tag__639276557962063929" := #enabled AND "ROLL_IO".Output[16, 7];
       "Tag__639276557962123762" := #enabled AND "ROLL_IO".Output[17, 0];
       "Tag__639276557962173628" := #enabled AND "ROLL_IO".Output[17, 1];
       "Tag__639276557962233470" := #enabled AND "ROLL_IO".Output[17, 2];
       "Tag__639276557962293353" := #enabled AND "ROLL_IO".Output[17, 3];
       "Tag__639276557962353158" := #enabled AND "ROLL_IO".Output[17, 4];
       "Tag__639276557962403014" := #enabled AND "ROLL_IO".Output[17, 5];
       "Tag__639276557962462907" := #enabled AND "ROLL_IO".Output[17, 6];
       "Tag__639276557962512720" := #enabled AND "ROLL_IO".Output[17, 7];
       "Tag__639276557962572561" := #enabled AND "ROLL_IO".Output[18, 0];
       "Tag__639276557962632401" := #enabled AND "ROLL_IO".Output[18, 1];
       "Tag__639276557962682267" := #enabled AND "ROLL_IO".Output[18, 2];
       "Tag__639276557962742107" := #enabled AND "ROLL_IO".Output[18, 3];
       "Tag__639276557962791974" := #enabled AND "ROLL_IO".Output[18, 4];
       "Tag__639276557962851816" := #enabled AND "ROLL_IO".Output[18, 5];
       "Tag__639276557962911653" := #enabled AND "ROLL_IO".Output[18, 6];
       "Tag__639276557962961520" := #enabled AND "ROLL_IO".Output[18, 7];
       "Tag__639276557963021363" := #enabled AND "ROLL_IO".Output[19, 0];
       "Tag__639276557963071237" := #enabled AND "ROLL_IO".Output[19, 1];
       "Tag__639276557963121101" := #enabled AND "ROLL_IO".Output[19, 2];
       "Tag__639276557963181309" := #enabled AND "ROLL_IO".Output[19, 3];
       "Tag__639276557963240774" := #enabled AND "ROLL_IO".Output[19, 4];
       "Tag__639276557963290937" := #enabled AND "ROLL_IO".Output[19, 5];
       "Tag__639276557963360463" := #enabled AND "ROLL_IO".Output[19, 6];
       "Tag__639276557963420293" := #enabled AND "ROLL_IO".Output[19, 7];
       "Tag__639276557963480133" := #enabled AND "ROLL_IO".Output[20, 0];
       "Tag__639276557963530002" := #enabled AND "ROLL_IO".Output[20, 1];
       "Tag__639276557963579865" := #enabled AND "ROLL_IO".Output[20, 2];
       "Tag__639276557963639838" := #enabled AND "ROLL_IO".Output[20, 3];
       "Tag__639276557963699546" := #enabled AND "ROLL_IO".Output[20, 4];
       "Tag__639276557963749412" := #enabled AND "ROLL_IO".Output[20, 5];
       "Tag__639276557963799286" := #enabled AND "ROLL_IO".Output[20, 6];
       "Tag__639276557963859119" := #enabled AND "ROLL_IO".Output[20, 7];
       "Tag__639276557963908985" := #enabled AND "ROLL_IO".Output[21, 0];
       "Tag__639276557963968826" := #enabled AND "ROLL_IO".Output[21, 1];
       "Tag__639276557964018692" := #enabled AND "ROLL_IO".Output[21, 2];
       "Tag__639276557964068878" := #enabled AND "ROLL_IO".Output[21, 3];
       "Tag__639276557964128400" := #enabled AND "ROLL_IO".Output[21, 4];
       "Tag__639276557964188239" := #enabled AND "ROLL_IO".Output[21, 5];
       "Tag__639276557964248077" := #enabled AND "ROLL_IO".Output[21, 6];
       "Tag__639276557964298411" := #enabled AND "ROLL_IO".Output[21, 7];
       "Tag__639276557964357785" := #enabled AND "ROLL_IO".Output[22, 0];
       "Tag__639276557964417947" := #enabled AND "ROLL_IO".Output[22, 1];
       "Tag__639276557964477465" := #enabled AND "ROLL_IO".Output[22, 2];
       "Tag__639276557964527497" := #enabled AND "ROLL_IO".Output[22, 3];
       "Tag__639276557964587312" := #enabled AND "ROLL_IO".Output[22, 4];
       "Tag__639276557964637070" := #enabled AND "ROLL_IO".Output[22, 5];
       "Tag__639276557964697149" := #enabled AND "ROLL_IO".Output[22, 6];
       "Tag__639276557964746745" := #enabled AND "ROLL_IO".Output[22, 7];
       "Tag__639276557964816574" := #enabled AND "ROLL_IO".Output[23, 0];
       "Tag__639276557964876412" := #enabled AND "ROLL_IO".Output[23, 1];
       "Tag__639276557964936239" := #enabled AND "ROLL_IO".Output[23, 2];
       "Tag__639276557964986111" := #enabled AND "ROLL_IO".Output[23, 3];
       "Tag__639276557965046275" := #enabled AND "ROLL_IO".Output[23, 4];
       "Tag__639276557965095821" := #enabled AND "ROLL_IO".Output[23, 5];
       "Tag__639276557965155664" := #enabled AND "ROLL_IO".Output[23, 6];
       "Tag__639276557965205527" := #enabled AND "ROLL_IO".Output[23, 7];
       "Tag__639276557965265365" := #enabled AND "ROLL_IO".Output[24, 0];
       "Tag__639276557965325265" := #enabled AND "ROLL_IO".Output[24, 1];
       "Tag__639276557965375063" := #enabled AND "ROLL_IO".Output[24, 2];
       "Tag__639276557965434904" := #enabled AND "ROLL_IO".Output[24, 3];
       "Tag__639276557965484769" := #enabled AND "ROLL_IO".Output[24, 4];
       "Tag__639276557965544610" := #enabled AND "ROLL_IO".Output[24, 5];
       "Tag__639276557965604458" := #enabled AND "ROLL_IO".Output[24, 6];
       "Tag__639276557965654714" := #enabled AND "ROLL_IO".Output[24, 7];
       "Tag__639276557965714166" := #enabled AND "ROLL_IO".Output[25, 0];
       "Tag__639276557965774008" := #enabled AND "ROLL_IO".Output[25, 1];
       "Tag__639276557965834033" := #enabled AND "ROLL_IO".Output[25, 2];
       "Tag__639276557965893680" := #enabled AND "ROLL_IO".Output[25, 3];
       "Tag__639276557965953516" := #enabled AND "ROLL_IO".Output[25, 4];
       "Tag__639276557966003383" := #enabled AND "ROLL_IO".Output[25, 5];
       "Tag__639276557966063222" := #enabled AND "ROLL_IO".Output[25, 6];
       "Tag__639276557966113089" := #enabled AND "ROLL_IO".Output[25, 7];
   END_IF;
END_FUNCTION
